(****************************************************************************************************<br>
© Syntegon Group.<br>
All rights reserved, also regarding any disposal, exploitation, reproduction, editing, distribution,<br>
as well as in the event of applications for industrial property rights.<br>
*****************************************************************************************************<br>
DESCRIPTION:<br>
TcUnit test suite of a parameter FB's m_Cycle (ADR 0017), on SynConfig._FB_ConfigConveyor: the program values<br>
while no set is active, a staged set taken over, waiting while the application does not allow it, rejected on<br>
another active version or when invalid, and a reset back to the program values. The tests write vo_Config's<br>
stStaging and stStaged as the gateway does over ADS.<br>
*****************************************************************************************************<br>
VERSION         ¦ DATE       ¦ NAME      ¦ CHANGE<br>
Syn_Config 2.0.0 ¦ 2026-11-11 ¦ J.Willner ¦ Unit tests<br>
Syn_Config 2.3.0 ¦ 2026-11-14 ¦ J.Willner ¦ The lifecycle of every parameter FB type<br>
****************************************************************************************************)
FUNCTION_BLOCK _FB_TestConfigStaging EXTENDS TcUnit.FB_TestSuite

m_ProgramValuesWithoutSet();
m_StagedSetTakenOver();
m_StagedSetWaitsUntilAllowed();
m_StagedSetOnOtherVersionRejected();
m_ResetReturnsToProgramValues();
m_InvalidProductTypesRejected();
m_EveryTypeRunsTheLifecycle();

(****************************************************************************************************<br>
© Syntegon Group.<br>
All rights reserved, also regarding any disposal, exploitation, reproduction, editing, distribution,<br>
as well as in the event of applications for industrial property rights.<br>
*****************************************************************************************************<br>
DESCRIPTION:<br>
Every parameter FB type runs the same staging lifecycle as the conveyor: a set staged on version 0 is taken over<br>
as version 1, a set staged on version 0 again is rejected (version 1 is active), and a reset returns to the<br>
program values under version 0. The machine FB's recipe has its own suite (_FB_TestConfigMachine).<br>
****************************************************************************************************)
METHOD PRIVATE m_EveryTypeRunsTheLifecycle
VAR_INST
	fb_TempDelta						: SynConfig._FB_ConfigDelta;
	TempDeltaDefault					: SynConfig.ST_ConfigDeltaParam;
	TempDeltaStaged						: SynConfig.ST_ConfigDeltaParam;
	TempDeltaSet						: SynConfig.ST_ConfigDeltaSet;
	fb_TempGantry						: SynConfig._FB_ConfigXtsGantry;
	TempGantryDefault					: SynConfig.ST_ConfigXtsGantryParam;
	TempGantryStaged					: SynConfig.ST_ConfigXtsGantryParam;
	TempGantrySet						: SynConfig.ST_ConfigXtsGantrySet;
	fb_TempLoop							: SynConfig._FB_ConfigXtsLoop;
	TempLoopDefault						: SynConfig.ST_ConfigXtsLoopParam;
	TempLoopStaged						: SynConfig.ST_ConfigXtsLoopParam;
	TempLoopSet							: SynConfig.ST_ConfigXtsLoopSet;
	fb_TempCartesian					: SynConfig._FB_ConfigCartesian;
	TempCartesianDefault				: SynConfig.ST_ConfigCartesianParam;
	TempCartesianStaged					: SynConfig.ST_ConfigCartesianParam;
	TempCartesianSet					: SynConfig.ST_ConfigCartesianSet;
	fb_TempVision						: SynConfig._FB_ConfigVision;
	TempVisionDefault					: SynConfig.ST_ConfigBodyComponentParam;
	TempVisionStaged					: SynConfig.ST_ConfigBodyComponentParam;
	TempVisionSet						: SynConfig.ST_ConfigBodyComponentSet;
	b_TempDone							: BOOL;	// the test ran
END_VAR
VAR
	b_TempChanged						: ARRAY[1..5, 1..3] OF BOOL;	// per type and step: m_Cycle's result
	e_TempResult						: ARRAY[1..5, 1..3] OF SynConfig.E_ConfigResult;	// per type and step: stStatus.eResult
	udn_TempVersion						: ARRAY[1..5, 1..3] OF UDINT;	// [-] per type and step: stStatus.nActiveVersion
	lr_TempX							: ARRAY[1..5, 1..3] OF LREAL;	// [mm] per type and step: X of the effective pose
	TempPose							: ST_VisuPose;
	un_TempStep							: UINT;	// [-] 1 = take-over, 2 = stale version, 3 = reset
	un_TempType							: UINT;
	p_TempDelta							: POINTER TO SynConfig.ST_ConfigDeltaParam;
	p_TempGantry						: POINTER TO SynConfig.ST_ConfigXtsGantryParam;
	p_TempLoop							: POINTER TO SynConfig.ST_ConfigXtsLoopParam;
	p_TempCartesian						: POINTER TO SynConfig.ST_ConfigCartesianParam;
	p_TempVision						: POINTER TO SynConfig.ST_ConfigBodyComponentParam;
END_VAR
VAR CONSTANT
	str_TYPE_NAMES						: ARRAY[1..5] OF STRING(20) := ['Delta', 'XTS gantry', 'XTS loop', 'Cartesian', 'Vision'];
END_VAR
TEST('ConfigEveryTypeRunsTheLifecycle');
IF b_TempDone THEN
	RETURN;
END_IF
b_TempDone := TRUE;


(****************************************************************************************************
THREE STEPS PER TYPE: TAKE-OVER, STALE VERSION, RESET
****************************************************************************************************)
(* Delta *)
TempDeltaDefault.stPose.fX := 100;
TempDeltaStaged.stPose.fX := 250;
p_TempDelta := ADR(fb_TempDelta.vo_Config.stStaged);
FOR un_TempStep := 1 TO 3 DO
	p_TempDelta^ := TempDeltaStaged;
	_FC_TestConfigStage(vi_p_Staging := ADR(fb_TempDelta.vo_Config.stStaging), vi_udn_BaseVersion := 0,
		vi_udn_StageId := UINT_TO_UDINT(un_TempStep), vi_b_Reset := un_TempStep = 3);
	b_TempChanged[1, un_TempStep] := fb_TempDelta.m_Cycle(vio_Default := TempDeltaDefault, vio_Set := TempDeltaSet,
		vi_b_ApplyAllowed := TRUE);
	e_TempResult[1, un_TempStep] := fb_TempDelta.vo_Config.stStatus.eResult;
	udn_TempVersion[1, un_TempStep] := fb_TempDelta.vo_Config.stStatus.nActiveVersion;
	TempPose := fb_TempDelta.m_Pose();
	lr_TempX[1, un_TempStep] := TempPose.fX;
END_FOR

(* XTS gantry: a track needs a module *)
TempGantryDefault.stPose.fX := 100;
TempGantryStaged.stPose.fX := 250;
TempGantryStaged.nModuleCount := 1;
TempGantryStaged.aModules[0].fLength := 250;
p_TempGantry := ADR(fb_TempGantry.vo_Config.stStaged);
FOR un_TempStep := 1 TO 3 DO
	p_TempGantry^ := TempGantryStaged;
	_FC_TestConfigStage(vi_p_Staging := ADR(fb_TempGantry.vo_Config.stStaging), vi_udn_BaseVersion := 0,
		vi_udn_StageId := UINT_TO_UDINT(un_TempStep), vi_b_Reset := un_TempStep = 3);
	b_TempChanged[2, un_TempStep] := fb_TempGantry.m_Cycle(vio_Default := TempGantryDefault, vio_Set := TempGantrySet,
		vi_b_ApplyAllowed := TRUE);
	e_TempResult[2, un_TempStep] := fb_TempGantry.vo_Config.stStatus.eResult;
	udn_TempVersion[2, un_TempStep] := fb_TempGantry.vo_Config.stStatus.nActiveVersion;
	TempPose := fb_TempGantry.m_Pose();
	lr_TempX[2, un_TempStep] := TempPose.fX;
END_FOR

(* XTS loop: a track needs a module *)
TempLoopDefault.stPose.fX := 100;
TempLoopStaged.stPose.fX := 250;
TempLoopStaged.nModuleCount := 1;
TempLoopStaged.aModules[0].fLength := 250;
p_TempLoop := ADR(fb_TempLoop.vo_Config.stStaged);
FOR un_TempStep := 1 TO 3 DO
	p_TempLoop^ := TempLoopStaged;
	_FC_TestConfigStage(vi_p_Staging := ADR(fb_TempLoop.vo_Config.stStaging), vi_udn_BaseVersion := 0,
		vi_udn_StageId := UINT_TO_UDINT(un_TempStep), vi_b_Reset := un_TempStep = 3);
	b_TempChanged[3, un_TempStep] := fb_TempLoop.m_Cycle(vio_Default := TempLoopDefault, vio_Set := TempLoopSet,
		vi_b_ApplyAllowed := TRUE);
	e_TempResult[3, un_TempStep] := fb_TempLoop.vo_Config.stStatus.eResult;
	udn_TempVersion[3, un_TempStep] := fb_TempLoop.vo_Config.stStatus.nActiveVersion;
	TempPose := fb_TempLoop.m_Pose();
	lr_TempX[3, un_TempStep] := TempPose.fX;
END_FOR

(* Cartesian *)
TempCartesianDefault.stPose.fX := 100;
TempCartesianStaged.stPose.fX := 250;
p_TempCartesian := ADR(fb_TempCartesian.vo_Config.stStaged);
FOR un_TempStep := 1 TO 3 DO
	p_TempCartesian^ := TempCartesianStaged;
	_FC_TestConfigStage(vi_p_Staging := ADR(fb_TempCartesian.vo_Config.stStaging), vi_udn_BaseVersion := 0,
		vi_udn_StageId := UINT_TO_UDINT(un_TempStep), vi_b_Reset := un_TempStep = 3);
	b_TempChanged[4, un_TempStep] := fb_TempCartesian.m_Cycle(vio_Default := TempCartesianDefault,
		vio_Set := TempCartesianSet, vi_b_ApplyAllowed := TRUE);
	e_TempResult[4, un_TempStep] := fb_TempCartesian.vo_Config.stStatus.eResult;
	udn_TempVersion[4, un_TempStep] := fb_TempCartesian.vo_Config.stStatus.nActiveVersion;
	TempPose := fb_TempCartesian.m_Pose();
	lr_TempX[4, un_TempStep] := TempPose.fX;
END_FOR

(* Vision system, for the body components *)
TempVisionDefault.stPose.fX := 100;
TempVisionStaged.stPose.fX := 250;
p_TempVision := ADR(fb_TempVision.vo_Config.stStaged);
FOR un_TempStep := 1 TO 3 DO
	p_TempVision^ := TempVisionStaged;
	_FC_TestConfigStage(vi_p_Staging := ADR(fb_TempVision.vo_Config.stStaging), vi_udn_BaseVersion := 0,
		vi_udn_StageId := UINT_TO_UDINT(un_TempStep), vi_b_Reset := un_TempStep = 3);
	b_TempChanged[5, un_TempStep] := fb_TempVision.m_Cycle(vio_Default := TempVisionDefault, vio_Set := TempVisionSet,
		vi_b_ApplyAllowed := TRUE);
	e_TempResult[5, un_TempStep] := fb_TempVision.vo_Config.stStatus.eResult;
	udn_TempVersion[5, un_TempStep] := fb_TempVision.vo_Config.stStatus.nActiveVersion;
	TempPose := fb_TempVision.m_Pose();
	lr_TempX[5, un_TempStep] := TempPose.fX;
END_FOR


(****************************************************************************************************
THE SAME RESULTS FOR EVERY TYPE
****************************************************************************************************)
FOR un_TempType := 1 TO 5 DO
	AssertTrue(Condition := b_TempChanged[un_TempType, 1], Message := CONCAT(str_TYPE_NAMES[un_TempType], ': taken over'));
	AssertEquals_UDINT(Expected := 1, Actual := udn_TempVersion[un_TempType, 1],
		Message := CONCAT(str_TYPE_NAMES[un_TempType], ': version 1 active'));
	AssertEquals_LREAL(Expected := 250, Actual := lr_TempX[un_TempType, 1], Delta := 0.001,
		Message := CONCAT(str_TYPE_NAMES[un_TempType], ': staged pose effective'));
	AssertFalse(Condition := b_TempChanged[un_TempType, 2],
		Message := CONCAT(str_TYPE_NAMES[un_TempType], ': stale version not taken over'));
	AssertTrue(Condition := e_TempResult[un_TempType, 2] = SynConfig.E_ConfigResult.REJECTED,
		Message := CONCAT(str_TYPE_NAMES[un_TempType], ': stale version rejected'));
	AssertEquals_UDINT(Expected := 1, Actual := udn_TempVersion[un_TempType, 2],
		Message := CONCAT(str_TYPE_NAMES[un_TempType], ': version 1 stays'));
	AssertTrue(Condition := b_TempChanged[un_TempType, 3], Message := CONCAT(str_TYPE_NAMES[un_TempType], ': reset'));
	AssertEquals_UDINT(Expected := 0, Actual := udn_TempVersion[un_TempType, 3],
		Message := CONCAT(str_TYPE_NAMES[un_TempType], ': version 0 after the reset'));
	AssertEquals_LREAL(Expected := 100, Actual := lr_TempX[un_TempType, 3], Delta := 0.001,
		Message := CONCAT(str_TYPE_NAMES[un_TempType], ': program pose again'));
END_FOR

TEST_FINISHED();
END_METHOD

(****************************************************************************************************<br>
© Syntegon Group.<br>
All rights reserved, also regarding any disposal, exploitation, reproduction, editing, distribution,<br>
as well as in the event of applications for industrial property rights.<br>
*****************************************************************************************************<br>
DESCRIPTION:<br>
A conveyor set is rejected with the reason when a product type has no number, a number is used twice or there<br>
are more product types than the list holds; the active set stays as it was.<br>
****************************************************************************************************)
METHOD PRIVATE m_InvalidProductTypesRejected
VAR_INST
	fb_TempParam						: SynConfig._FB_ConfigConveyor;
	TempDefault							: SynConfig.ST_ConfigConveyorParam;
	TempSet								: SynConfig.ST_ConfigConveyorSet;
	b_TempDone							: BOOL;	// the test ran
END_VAR
VAR
	TempStaged							: SynConfig.ST_ConfigConveyorParam;
END_VAR
TEST('ConfigInvalidProductTypesRejected');
IF b_TempDone THEN
	RETURN;
END_IF
b_TempDone := TRUE;

TempDefault := m_ValidSet(vi_lr_X := 100);

(* A product type without a number. *)
TempStaged := m_ValidSet(vi_lr_X := 250);
TempStaged.aProductTypes[1].nId := 0;
m_Stage(vio_Param := fb_TempParam, vio_Staged := TempStaged, vi_udn_BaseVersion := 0, vi_udn_StageId := 1);
AssertFalse(Condition := fb_TempParam.m_Cycle(vio_Default := TempDefault, vio_Set := TempSet, vi_b_ApplyAllowed := TRUE),
	Message := 'type without a number: not taken over');
AssertTrue(Condition := fb_TempParam.vo_Config.stStatus.eResult = SynConfig.E_ConfigResult.REJECTED, Message := 'rejected');
AssertEquals_STRING(Expected := 'A product type without a number', Actual := fb_TempParam.vo_Config.stStatus.sMessage,
	Message := 'reason: no number');

(* A number used twice. *)
TempStaged := m_ValidSet(vi_lr_X := 250);
TempStaged.aProductTypes[0].nId := 3;
TempStaged.aProductTypes[1].nId := 3;
m_Stage(vio_Param := fb_TempParam, vio_Staged := TempStaged, vi_udn_BaseVersion := 0, vi_udn_StageId := 2);
AssertFalse(Condition := fb_TempParam.m_Cycle(vio_Default := TempDefault, vio_Set := TempSet, vi_b_ApplyAllowed := TRUE),
	Message := 'number twice: not taken over');
AssertEquals_STRING(Expected := 'Product type 3 is defined twice', Actual := fb_TempParam.vo_Config.stStatus.sMessage,
	Message := 'reason: defined twice');

(* More product types than the list holds. *)
TempStaged := m_ValidSet(vi_lr_X := 250);
TempStaged.nProductTypeCount := VISU_GlobalConst_Param.VISU_un_MAX_PRODUCT_TYPES + 1;
m_Stage(vio_Param := fb_TempParam, vio_Staged := TempStaged, vi_udn_BaseVersion := 0, vi_udn_StageId := 3);
AssertFalse(Condition := fb_TempParam.m_Cycle(vio_Default := TempDefault, vio_Set := TempSet, vi_b_ApplyAllowed := TRUE),
	Message := 'too many types: not taken over');
AssertEquals_STRING(Expected := CONCAT('More than ', CONCAT(UINT_TO_STRING(VISU_GlobalConst_Param.VISU_un_MAX_PRODUCT_TYPES),
	' product types')), Actual := fb_TempParam.vo_Config.stStatus.sMessage, Message := 'reason: too many');
AssertEquals_UDINT(Expected := 3, Actual := fb_TempParam.vo_Config.stStatus.nHandledStageId, Message := 'last stage id handled');

AssertFalse(Condition := TempSet.bValid, Message := 'still no active set');
AssertEquals_LREAL(Expected := 100, Actual := fb_TempParam.vo_Config.stActive.stPose.fX, Delta := 0.001,
	Message := 'program values still effective');

TEST_FINISHED();
END_METHOD

(****************************************************************************************************<br>
© Syntegon Group.<br>
All rights reserved, also regarding any disposal, exploitation, reproduction, editing, distribution,<br>
as well as in the event of applications for industrial property rights.<br>
*****************************************************************************************************<br>
DESCRIPTION:<br>
Without an active set the program values are effective, under version 0, and nothing has been handled.<br>
****************************************************************************************************)
METHOD PRIVATE m_ProgramValuesWithoutSet
VAR_INST
	fb_TempParam						: SynConfig._FB_ConfigConveyor;
	TempDefault							: SynConfig.ST_ConfigConveyorParam;
	TempSet								: SynConfig.ST_ConfigConveyorSet;
	b_TempDone							: BOOL;	// the test ran
END_VAR
VAR
	TempPose							: ST_VisuPose;
END_VAR
TEST('ConfigProgramValuesWithoutSet');
IF b_TempDone THEN
	RETURN;
END_IF
b_TempDone := TRUE;

TempDefault := m_ValidSet(vi_lr_X := 100);
AssertFalse(Condition := fb_TempParam.m_Cycle(vio_Default := TempDefault, vio_Set := TempSet, vi_b_ApplyAllowed := TRUE),
	Message := 'nothing staged: no change');
TempPose := fb_TempParam.m_Pose();
AssertEquals_LREAL(Expected := 100, Actual := TempPose.fX, Delta := 0.001, Message := 'program pose effective');
AssertEquals_UINT(Expected := 2, Actual := fb_TempParam.vo_Config.stActive.nProductTypeCount, Message := 'program product types effective');
AssertEquals_UDINT(Expected := 0, Actual := fb_TempParam.vo_Config.stStatus.nActiveVersion, Message := 'version 0: program values');
AssertTrue(Condition := fb_TempParam.vo_Config.stStatus.eResult = SynConfig.E_ConfigResult.NONE, Message := 'nothing handled');

TEST_FINISHED();
END_METHOD

(****************************************************************************************************<br>
© Syntegon Group.<br>
All rights reserved, also regarding any disposal, exploitation, reproduction, editing, distribution,<br>
as well as in the event of applications for industrial property rights.<br>
*****************************************************************************************************<br>
DESCRIPTION:<br>
A reset makes the active set invalid at once (also while a take-over is not allowed): the program values apply<br>
under version 0. Versions never repeat: the next set taken over gets version 2, not 1.<br>
****************************************************************************************************)
METHOD PRIVATE m_ResetReturnsToProgramValues
VAR_INST
	fb_TempParam						: SynConfig._FB_ConfigConveyor;
	TempDefault							: SynConfig.ST_ConfigConveyorParam;
	TempSet								: SynConfig.ST_ConfigConveyorSet;
	b_TempDone							: BOOL;	// the test ran
END_VAR
VAR
	TempStaged							: SynConfig.ST_ConfigConveyorParam;
END_VAR
TEST('ConfigResetReturnsToProgramValues');
IF b_TempDone THEN
	RETURN;
END_IF
b_TempDone := TRUE;

TempDefault := m_ValidSet(vi_lr_X := 100);
TempStaged := m_ValidSet(vi_lr_X := 250);
m_Stage(vio_Param := fb_TempParam, vio_Staged := TempStaged, vi_udn_BaseVersion := 0, vi_udn_StageId := 1);
fb_TempParam.m_Cycle(vio_Default := TempDefault, vio_Set := TempSet, vi_b_ApplyAllowed := TRUE);
AssertEquals_UDINT(Expected := 1, Actual := fb_TempParam.vo_Config.stStatus.nActiveVersion, Message := 'version 1 active');

_FC_TestConfigStage(vi_p_Staging := ADR(fb_TempParam.vo_Config.stStaging), vi_udn_BaseVersion := 1, vi_udn_StageId := 2,
	vi_b_Reset := TRUE);
AssertTrue(Condition := fb_TempParam.m_Cycle(vio_Default := TempDefault, vio_Set := TempSet, vi_b_ApplyAllowed := FALSE),
	Message := 'reset handled, even while not allowed');
AssertFalse(Condition := TempSet.bValid, Message := 'active set invalid');
AssertEquals_UDINT(Expected := 0, Actual := fb_TempParam.vo_Config.stStatus.nActiveVersion, Message := 'version 0');
AssertEquals_LREAL(Expected := 100, Actual := fb_TempParam.vo_Config.stActive.stPose.fX, Delta := 0.001,
	Message := 'program values effective again');
AssertTrue(Condition := fb_TempParam.vo_Config.stStatus.eResult = SynConfig.E_ConfigResult.APPLIED, Message := 'reset applied');
AssertEquals_UDINT(Expected := 2, Actual := fb_TempParam.vo_Config.stStatus.nHandledStageId, Message := 'stage id handled');
AssertFalse(Condition := fb_TempParam.vo_Config.stStaging.bReset, Message := 'reset flag cleared');

m_Stage(vio_Param := fb_TempParam, vio_Staged := TempStaged, vi_udn_BaseVersion := 0, vi_udn_StageId := 3);
fb_TempParam.m_Cycle(vio_Default := TempDefault, vio_Set := TempSet, vi_b_ApplyAllowed := TRUE);
AssertEquals_UDINT(Expected := 2, Actual := fb_TempParam.vo_Config.stStatus.nActiveVersion, Message := 'next set gets version 2');

TEST_FINISHED();
END_METHOD

(****************************************************************************************************<br>
© Syntegon Group.<br>
All rights reserved, also regarding any disposal, exploitation, reproduction, editing, distribution,<br>
as well as in the event of applications for industrial property rights.<br>
*****************************************************************************************************<br>
DESCRIPTION:<br>
Stages a set on a conveyor's parameter FB as the gateway does: the set into vo_Config.stStaged, then stStaging<br>
(_FC_TestConfigStage). The FB handles it in its next m_Cycle.<br>
****************************************************************************************************)
METHOD PRIVATE m_Stage : BOOL
VAR_IN_OUT
	vio_Param							: SynConfig._FB_ConfigConveyor;	// the parameter FB under test
END_VAR
VAR_IN_OUT CONSTANT
	vio_Staged							: SynConfig.ST_ConfigConveyorParam;	// the set to stage
END_VAR
VAR_INPUT
	vi_udn_BaseVersion					: UDINT;	// [-] active version the set is based on
	vi_udn_StageId						: UDINT;	// [-] the gateway's id of this staging
END_VAR
VAR
	p_TempStaged						: POINTER TO SynConfig.ST_ConfigConveyorParam;
END_VAR
p_TempStaged := ADR(vio_Param.vo_Config.stStaged);
p_TempStaged^ := vio_Staged;
m_Stage := _FC_TestConfigStage(vi_p_Staging := ADR(vio_Param.vo_Config.stStaging), vi_udn_BaseVersion := vi_udn_BaseVersion,
	vi_udn_StageId := vi_udn_StageId, vi_b_Reset := FALSE);
END_METHOD

(****************************************************************************************************<br>
© Syntegon Group.<br>
All rights reserved, also regarding any disposal, exploitation, reproduction, editing, distribution,<br>
as well as in the event of applications for industrial property rights.<br>
*****************************************************************************************************<br>
DESCRIPTION:<br>
A set staged on another version than the active one is rejected with the reason, even while a take-over is<br>
allowed: someone else changed the set since the configurator read it.<br>
****************************************************************************************************)
METHOD PRIVATE m_StagedSetOnOtherVersionRejected
VAR_INST
	fb_TempParam						: SynConfig._FB_ConfigConveyor;
	TempDefault							: SynConfig.ST_ConfigConveyorParam;
	TempSet								: SynConfig.ST_ConfigConveyorSet;
	b_TempDone							: BOOL;	// the test ran
END_VAR
VAR
	TempStaged							: SynConfig.ST_ConfigConveyorParam;
END_VAR
TEST('ConfigStagedSetOnOtherVersionRejected');
IF b_TempDone THEN
	RETURN;
END_IF
b_TempDone := TRUE;

TempDefault := m_ValidSet(vi_lr_X := 100);
TempStaged := m_ValidSet(vi_lr_X := 250);
m_Stage(vio_Param := fb_TempParam, vio_Staged := TempStaged, vi_udn_BaseVersion := 5, vi_udn_StageId := 9);

AssertFalse(Condition := fb_TempParam.m_Cycle(vio_Default := TempDefault, vio_Set := TempSet, vi_b_ApplyAllowed := TRUE),
	Message := 'not taken over');
AssertTrue(Condition := fb_TempParam.vo_Config.stStatus.eResult = SynConfig.E_ConfigResult.REJECTED, Message := 'rejected');
AssertEquals_STRING(Expected := 'Based on version 5, but version 0 is active', Actual := fb_TempParam.vo_Config.stStatus.sMessage,
	Message := 'the reason');
AssertEquals_UDINT(Expected := 9, Actual := fb_TempParam.vo_Config.stStatus.nHandledStageId, Message := 'stage id handled');
AssertFalse(Condition := fb_TempParam.vo_Config.stStaging.bStaged, Message := 'staged flag cleared');
AssertFalse(Condition := TempSet.bValid, Message := 'no active set');

TEST_FINISHED();
END_METHOD

(****************************************************************************************************<br>
© Syntegon Group.<br>
All rights reserved, also regarding any disposal, exploitation, reproduction, editing, distribution,<br>
as well as in the event of applications for industrial property rights.<br>
*****************************************************************************************************<br>
DESCRIPTION:<br>
A set staged on the active version is taken over while the application allows it: it becomes the active set<br>
under version 1 and the effective values, the status names the stage id as applied and the flags are cleared.<br>
****************************************************************************************************)
METHOD PRIVATE m_StagedSetTakenOver
VAR_INST
	fb_TempParam						: SynConfig._FB_ConfigConveyor;
	TempDefault							: SynConfig.ST_ConfigConveyorParam;
	TempSet								: SynConfig.ST_ConfigConveyorSet;
	b_TempDone							: BOOL;	// the test ran
END_VAR
VAR
	TempPose							: ST_VisuPose;
	TempStaged							: SynConfig.ST_ConfigConveyorParam;
END_VAR
TEST('ConfigStagedSetTakenOver');
IF b_TempDone THEN
	RETURN;
END_IF
b_TempDone := TRUE;

TempDefault := m_ValidSet(vi_lr_X := 100);
TempStaged := m_ValidSet(vi_lr_X := 250);
m_Stage(vio_Param := fb_TempParam, vio_Staged := TempStaged, vi_udn_BaseVersion := 0, vi_udn_StageId := 7);

AssertTrue(Condition := fb_TempParam.m_Cycle(vio_Default := TempDefault, vio_Set := TempSet, vi_b_ApplyAllowed := TRUE),
	Message := 'set taken over');
AssertTrue(Condition := TempSet.bValid, Message := 'active set valid');
AssertEquals_UDINT(Expected := 1, Actual := TempSet.nVersion, Message := 'first version');
AssertEquals_UDINT(Expected := 1, Actual := fb_TempParam.vo_Config.stStatus.nActiveVersion, Message := 'status names the version');
AssertEquals_UDINT(Expected := 7, Actual := fb_TempParam.vo_Config.stStatus.nHandledStageId, Message := 'stage id handled');
AssertTrue(Condition := fb_TempParam.vo_Config.stStatus.eResult = SynConfig.E_ConfigResult.APPLIED, Message := 'applied');
AssertEquals_STRING(Expected := '', Actual := fb_TempParam.vo_Config.stStatus.sMessage, Message := 'no message');
AssertFalse(Condition := fb_TempParam.vo_Config.stStaging.bStaged, Message := 'staged flag cleared');
TempPose := fb_TempParam.m_Pose();
AssertEquals_LREAL(Expected := 250, Actual := TempPose.fX, Delta := 0.001, Message := 'staged pose effective');

AssertFalse(Condition := fb_TempParam.m_Cycle(vio_Default := TempDefault, vio_Set := TempSet, vi_b_ApplyAllowed := TRUE),
	Message := 'next cycle: no change');
AssertEquals_UDINT(Expected := 1, Actual := fb_TempParam.vo_Config.stStatus.nActiveVersion, Message := 'still version 1');

TEST_FINISHED();
END_METHOD

(****************************************************************************************************<br>
© Syntegon Group.<br>
All rights reserved, also regarding any disposal, exploitation, reproduction, editing, distribution,<br>
as well as in the event of applications for industrial property rights.<br>
*****************************************************************************************************<br>
DESCRIPTION:<br>
While the application does not allow a take-over the staged set waits (PENDING, still staged, the program values<br>
stay effective); it is taken over in the first cycle that allows it.<br>
****************************************************************************************************)
METHOD PRIVATE m_StagedSetWaitsUntilAllowed
VAR_INST
	fb_TempParam						: SynConfig._FB_ConfigConveyor;
	TempDefault							: SynConfig.ST_ConfigConveyorParam;
	TempSet								: SynConfig.ST_ConfigConveyorSet;
	b_TempDone							: BOOL;	// the test ran
END_VAR
VAR
	TempStaged							: SynConfig.ST_ConfigConveyorParam;
END_VAR
TEST('ConfigStagedSetWaitsUntilAllowed');
IF b_TempDone THEN
	RETURN;
END_IF
b_TempDone := TRUE;

TempDefault := m_ValidSet(vi_lr_X := 100);
TempStaged := m_ValidSet(vi_lr_X := 250);
m_Stage(vio_Param := fb_TempParam, vio_Staged := TempStaged, vi_udn_BaseVersion := 0, vi_udn_StageId := 3);

AssertFalse(Condition := fb_TempParam.m_Cycle(vio_Default := TempDefault, vio_Set := TempSet, vi_b_ApplyAllowed := FALSE),
	Message := 'not allowed: not taken over');
AssertTrue(Condition := fb_TempParam.vo_Config.stStatus.eResult = SynConfig.E_ConfigResult.PENDING, Message := 'pending');
AssertTrue(Condition := fb_TempParam.vo_Config.stStaging.bStaged, Message := 'still staged');
AssertFalse(Condition := TempSet.bValid, Message := 'no active set yet');
AssertEquals_LREAL(Expected := 100, Actual := fb_TempParam.vo_Config.stActive.stPose.fX, Delta := 0.001,
	Message := 'program values still effective');

AssertTrue(Condition := fb_TempParam.m_Cycle(vio_Default := TempDefault, vio_Set := TempSet, vi_b_ApplyAllowed := TRUE),
	Message := 'allowed: taken over');
AssertTrue(Condition := fb_TempParam.vo_Config.stStatus.eResult = SynConfig.E_ConfigResult.APPLIED, Message := 'applied');
AssertEquals_UDINT(Expected := 3, Actual := fb_TempParam.vo_Config.stStatus.nHandledStageId, Message := 'stage id handled');

TEST_FINISHED();
END_METHOD

(****************************************************************************************************<br>
© Syntegon Group.<br>
All rights reserved, also regarding any disposal, exploitation, reproduction, editing, distribution,<br>
as well as in the event of applications for industrial property rights.<br>
*****************************************************************************************************<br>
DESCRIPTION:<br>
A conveyor parameter set that can be taken over: the pose at X = vi_lr_X and two product types (1 and 2).<br>
****************************************************************************************************)
METHOD PRIVATE m_ValidSet : SynConfig.ST_ConfigConveyorParam
VAR_INPUT
	vi_lr_X								: LREAL;	// [mm] X of the pose, to tell sets apart
END_VAR
m_ValidSet.stPose.fX := vi_lr_X;
m_ValidSet.stOriginShift.fX := 50;
m_ValidSet.nProductTypeCount := 2;
m_ValidSet.aProductTypes[0].nId := 1;
m_ValidSet.aProductTypes[0].fLength := 120;
m_ValidSet.aProductTypes[0].fWidth := 80;
m_ValidSet.aProductTypes[0].fHeight := 40;
m_ValidSet.aProductTypes[0].eShape := E_VisuProductShape.BOX;
m_ValidSet.aProductTypes[1].nId := 2;
m_ValidSet.aProductTypes[1].fLength := 66;
m_ValidSet.aProductTypes[1].fWidth := 66;
m_ValidSet.aProductTypes[1].fHeight := 120;
m_ValidSet.aProductTypes[1].eShape := E_VisuProductShape.CYLINDER;
END_METHOD

END_FUNCTION_BLOCK

(* stored: Version 1.1.0.1
   POU _FB_TestConfigStaging: Id {4e682200-50f1-4b62-b8ee-93797b6552a3}, SpecialFunc None
   Method m_EveryTypeRunsTheLifecycle: Id {98d7e76b-db1d-4f02-9bf1-fe0eb3da25fc}
   Method m_InvalidProductTypesRejected: Id {5b5ed334-7115-4d9e-9594-25e6249f4a24}
   Method m_ProgramValuesWithoutSet: Id {1bc8d81c-74f6-41d8-a970-13ac87471f98}
   Method m_ResetReturnsToProgramValues: Id {6ed7f933-143f-4eb7-81ed-da42e795bd9b}
   Method m_Stage: Id {48432c50-6d91-4cca-a58b-d61e8c68e499}
   Method m_StagedSetOnOtherVersionRejected: Id {c6cdc518-4a54-429b-ad76-26e750b0444a}
   Method m_StagedSetTakenOver: Id {b7908878-aabf-4eae-b270-bed79057eaef}
   Method m_StagedSetWaitsUntilAllowed: Id {1329ac46-7b87-459b-b58c-78c66470069c}
   Method m_ValidSet: Id {57369c18-e466-45fb-a01b-f72ef93ea21f} *)
